// TIA Portal V21 export
// export: Created 2026-11-11T00:47:29.7188269Z, ExportSetting WithDefaults, DisplayName Totally Integrated Automation Portal, DisplayVersion V21 Update 3, DisplayName STEP 7 Professional, DisplayVersion V21 Update 3, DisplayName STEP 7 Safety, DisplayVersion V21, DisplayName Tech WebApplication, DisplayVersion V21, DisplayName WinCC Basic/Comfort/Advanced, DisplayVersion V21 Update 3, DisplayName WinCC Unified, DisplayVersion V21 Update 3
FUNCTION_BLOCK "FB_Fbd_ex114"   // FB126, FBD
{ S7_Optimized_Access := 'TRUE' }
VERSION : 0.1
// stored: AutoNumber true, IsIECCheckEnabled false, IsRetainMemResEnabled false, MemoryReserve 100, SetENOAutomatically false, UDAEnableTagReadback false
   VAR_INPUT
      v_prgflt_query : DWord;
      v_accflt_query : DWord;
   END_VAR
   VAR_OUTPUT
      v_ret_val : Int;
      v_prgflt_clr : DWord;
      v_accflt_clr : DWord;
   END_VAR
BEGIN

REGION Network 1: READ_ERR - Read out event status register
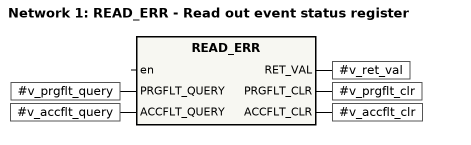
   #v_ret_val := READ_ERR(PRGFLT_QUERY := #v_prgflt_query,
                          ACCFLT_QUERY := #v_accflt_query,
                          PRGFLT_CLR => #v_prgflt_clr,
                          ACCFLT_CLR => #v_accflt_clr);
END_REGION
END_FUNCTION_BLOCK
